(* IEC 61131-3 sources: SortJet_MasterSPS_Aufbau.fbsproj/09_Station/Shuttle/Bewegung, 2 files *)

(* ---- Querfahrt_Shuttle_FB_V01_00_00.fb.st ---- *)
(* METADATA
{
	"v3Meta": {
		"objectGuid": "72dffa9c-0dea-4fd7-9820-5307a69ebe3d"
	}
}
*)
FUNCTION_BLOCK Querfahrt_Shuttle_FB_V01_00_00
VAR_INPUT

  // BOOLEAN
  bpAktivieren                           : BOOL; // Hinweis: Baustein aktivieren
  bpReset                                : BOOL; // BETRIEBSART: Fehler zuruecksetzen
  bpReferenz                        : BOOL;
  bpHandfahrenPlus                             : BOOL;
  bpHandfahrenMinus                            : BOOL;
  bpFreigabe                             : BOOL; // Sicherheitsfreigabe Regler darf Freigeben
  bpAutomatikAktiv                       : BOOL; // BETRIEBSART: Umschaltung der Geschwindigkeit
  bpVerfahreShuttle                      : BOOL; // Befehl zum Positionieren
  bpVerfahrfreigabe                      : BOOL; // Das entsprechende Shutte setzt die Verfahrfreigabe und überträgt es an die Verfahrkontrolle
  bpSofortStop                           : BOOL;
  bpQuittungAuftragsstatusZurueckgesetzt : BOOL; // Auftrag wurde zurueckgesetzt
  bpTeilnehmerErreichbar                 : BOOL;
  bpShuttleFaecherwagenSuche             : BOOL;
  bpLangsamfahrtNockenAktivieren         : BOOL;

  // WORD
  wpAuftragsTyp                          : WORD; // Bit 1 = Positionierauftrag mit Messgeschwindigkeit (RackSuche), aus dem Positionierauftrag (Vorabpositionierung)

  // REAL
  rpDestinationPosition                  : REAL; // ZielPosition
  rpMinPosSwEsEingrenzung                : REAL;
  rpMaxPosSwEsEingrenzung                : REAL;

  // POINTER
  ppAntriebsInformationen  : REFERENCE TO AntriebsInformationen; // Hinweis: Beinhaltet die Geschwindigkeiten / Rampen der einzelnen Shuttle

  // STRUKTUR
  stStationsNummern     : Station_ST;

END_VAR
VAR_OUTPUT

  // BOOLEAN
  bpDone                         : BOOL;
  bpFehler                       : BOOL;
  bpPositionierungAktiv          : BOOL;
  bpAntriebLaeuft                : BOOL;
  bpInReference                  : BOOL;
  bpAuftragsstatusZuruecksetzen  : BOOL := FALSE;
  bpAbbruchPositionierung        : BOOL := FALSE;

  // WORD
  wpFehlerNr     : Fehlerkonstanten_EN; // Exception- Handle: Fehlernummer

  // REAL
  rpAktPosition : REAL;
  rpAktSpeed    : REAL;

  // HARDWARE EINGAENGE
  in_bLeistungsschutzFremdluefter : BOOL;
  in_bEndschalterMax              : BOOL; // Oeffner (TRUE = frei), gemappt; zum Umrichter ueber Signal-Steuerwort Bit 9, wirkt nur bei Endschalterquelle SPS
  in_bEndschalterMin              : BOOL; // Oeffner (TRUE = frei), gemappt; zum Umrichter ueber Signal-Steuerwort Bit 10, wirkt nur bei Endschalterquelle SPS

END_VAR
VAR

  // BOOLEAN
  Antrieb : REFERENCE TO Rexroth_ctrlX_Drive_Eckelmann_MC_V01_02_02;

  // BOOLEAN
  blErsterZyklus                : BOOL := TRUE;
  blFreigabeGesetzt             : BOOL;
  blAlterStatus_Bewegung        : BOOL;

  // REAL
  rlAlterStatus_Position        : REAL;

  // STEPS
  STEP_Mov_Shuttle_W    : Steps_TE;
  schrittlReset         : STEPS_TE;
  steplReferenz         : STEPS_TE;

  // TIMER
  tonlWarteAufStop                      : TON; // EINSCHALTVERZOEGERUNG:
  tonlWarteAufReset                     : TON; // EINSCHALTVERZOEGERUNG:
  tofAntriebFreigabe                    : TOF; // AUSSCHALTVERZÖGERUNG
  tonlEndschalterFreifahren             : TON;
  tonlWarteSchrittEndschalterFreifahren : TON;
  toflHardwareEndschalterFrei           : TOF;
  tonlSafetyTimeout                     : TON;
  tonlFreigabe                          : TON;
  tonlAntriebNichtBetriebsbereit        : TON;
  tonlStatusMelden                      : TON;

  // TRIGGER
  rtlAutoAktiv : R_TRIG;

END_VAR

//-------------------------------------------------------------------------------------------------
// S T A R T - Initialisierung
//-------------------------------------------------------------------------------------------------
IF ( blErsterZyklus ) THEN

  IF ( __ISVALIDREF(ppAntriebsInformationen) ) THEN

    blErsterZyklus := FALSE;

    Antrieb REF= pgAntriebe[ppAntriebsInformationen.wAchsID];

    (* Hinweis:
       - Initialisierung Antriebsinformationen
    *)
    Antrieb.ppAntriebsInformationen REF= ppAntriebsInformationen;
    Antrieb.stStationsNummern := stStationsNummern;

    (* Hinweis:
       - Für die Zielpunktkontrolle muss im ersten Zyklus (und nach jeder Referenzierung) die Zielposition initialisiert werden
    *)
    Antrieb.rpZielPosition := Antrieb.rpIstPosition;

    (* Hinweis:
       - Antriebswerte vorinitialisieren
    *)
    Antrieb.rpGeschwindigkeit := ppAntriebsInformationen.rpHandGeschwindigkeit;
    Antrieb.rpBeschleunigung  := ppAntriebsInformationen.rpMaxBeschleunigung;
    Antrieb.rpVerzoegerung    := ppAntriebsInformationen.rpMaxVerzoegerung;
    Antrieb.rpRuckzeit        := ppAntriebsInformationen.rpMaxRuckzeit;

  ELSE
    RETURN;
  END_IF

END_IF

//-------------------------------------------------------------------------------------------------
// E N D E - Initialisierung
//-------------------------------------------------------------------------------------------------

// Endschalter zyklisch an den Antrieb geben, auch bei deaktivierter Bewegung
Antrieb.bpEndschalterMinExtern := in_bEndschalterMin;
Antrieb.bpEndschalterMaxExtern := in_bEndschalterMax;

//-------------------------------------------------------------------------------------------------
// DEAKTIVIEREN
//-------------------------------------------------------------------------------------------------
IF ( NOT bpAktivieren ) THEN

  bpDone                        := TRUE;
  bpAuftragsstatusZuruecksetzen := FALSE;
  bpAbbruchPositionierung       := FALSE;

  bpFehler   := FALSE;
  wpFehlerNr := cMELDUNG_NULL;

  Antrieb.bpFreigabe := FALSE;

  RETURN;

END_IF

//-------------------------------------------------------------------------------------------------
// S T A R T - Timer
//-------------------------------------------------------------------------------------------------

rtlAutoAktiv(CLK := bpAutomatikAktiv);

IF ( rtlAutoAktiv.Q ) THEN
  Antrieb.rpZielPosition := Antrieb.rpIstPosition;
END_IF

(* Hinweis:
   - Aktuell wird diese Einschaltverzoegerung nur bei Motoren mit Bremse benoetigt [Lenze]
     => Eingebunden bei den Handfunktionen
*)
tofAntriebFreigabe( IN := blFreigabeGesetzt AND Antrieb.bpReglerBereit  , PT := T#10S );

// *************************************************************************************************

//-------------------------------------------------------------------------------------------------
// S T A R T - Verfahrschrittketten zurücksetzen
//-------------------------------------------------------------------------------------------------

// *************************************************************************************************

IF (   bpVerfahrfreigabe
     AND bpAbbruchPositionierung
     AND bpQuittungAuftragsstatusZurueckgesetzt )
THEN
  bpAbbruchPositionierung := FALSE;
  bpAuftragsstatusZuruecksetzen := FALSE;
  bpQuittungAuftragsstatusZurueckgesetzt := FALSE;

  wSps2MmiStationsNummer     := stStationsNummern.NummerIntern;
  rSps2MmiPosition           := Antrieb.rpIstPosition;
  MsgToMmi(SB0_SPS_SHUTTLEVORABPOSITIONIERUNGREADY);

END_IF

//-------------------------------------------------------------------------------------------------
// S T A R T - BAUSTEINE AUFRUFEN
//-------------------------------------------------------------------------------------------------

//-------------------------------------------------------------------------------------------------
// S T A R T - BAUSTEINE AUFRUFEN
//-------------------------------------------------------------------------------------------------
Verfahren();
Handfunktionen();
Referenz();
Reset();
Meldungen();

//-------------------------------------------------------------------------------------------------
// E N D E - BAUSTEINE AUFRUFEN
//-------------------------------------------------------------------------------------------------
IF ( bpSofortStop OR NOT abgVerfahrfreigabeShuttle[stStationsNummern.NummerSPS] ) OR NOT bpFreigabe THEN
  Antrieb.bpFreigabe := FALSE;
END_IF

Antrieb.stStationsNummern            := stStationsNummern;

Antrieb.bpAktiviereLangsamfahrtNocke := bpLangsamfahrtNockenAktivieren;
Antrieb.rpMinSwEsEingrenzung         := rpMinPosSwEsEingrenzung;
Antrieb.rpMaxSwEsEingrenzung         := rpMaxPosSwEsEingrenzung;

// übergabe der aktuellen Position
rpAktPosition   := Antrieb.rpIstPosition;
rpAktSpeed      := Antrieb.rpIstGeschwindigkeit; // mm/s, mit Vorzeichen
bpInReference   := Antrieb.bpIstReferenziert;
bpAntriebLaeuft := Antrieb.bpAntrieblaeuft;

// STATUS AN MMI MELDEN
tonlStatusMelden(
                  IN := NOT tonlStatusMelden.Q,
                  PT := T#500MS
                );

// Neue MMI-Verbindung (Flanke, nur ein Zyklus) sofort melden, nicht nur im 500-ms-Takt
IF    (     tonlStatusMelden.Q
        AND (    ( ABS( Antrieb.rpIstPosition - rlAlterStatus_Position ) > 1.0 )
              OR ( Antrieb.bpAntrieblaeuft <> blAlterStatus_Bewegung ) ) )
   OR Job.rtlMmiOk.Q
THEN
  stStationUpdate.wStationsNummer       := stStationsNummern.NummerSPS;
  stStationUpdate.eUpdateTyp            := StationUpdateTyp_EN.POSITIONSAENDERUNG;
  stStationUpdate.wAnzahlWerte          := 2;
  stStationUpdate.astWerte[1].eDatenTyp := UpdateDatenTyp_EN.TYP_REAL;
  stStationUpdate.astWerte[1].rWert     := Antrieb.rpIstPosition;
  stStationUpdate.astWerte[2].eDatenTyp := UpdateDatenTyp_EN.TYP_BOOL;
  stStationUpdate.astWerte[2].bWert     := Antrieb.bpAntrieblaeuft;
  MsgToMmi( auftragsnr_w := SB0_SPS_STATION_UPDATE );

  rlAlterStatus_Position := Antrieb.rpIstPosition;
  blAlterStatus_Bewegung := Antrieb.bpAntrieblaeuft;
END_IF
END_FUNCTION_BLOCK

(* ---- Verfahrueberwachung_PRG.prg.st ---- *)
(* METADATA
{
	"v3Meta": {
		"objectGuid": "88539335-6d2a-4efd-8213-a5feda61f359"
	}
}
*)
PROGRAM Verfahrueberwachung_PRG
VAR

  // BOOLEAN
  ablKonfiguriert                           : ARRAY[cERSTES_SHUTTLE..cLETZTES_TRANSFERSHUTTLE] OF BOOL; // Shuttle / Transfershuttle ist in dieser Anlage vorhanden
  ablShuttleInParkpos                       : ARRAY[cERSTES_SHUTTLE..cLETZTES_TRANSFERSHUTTLE] OF BOOL;
  ablShuttleStehtOhnePositionsveraenderung  : ARRAY[cERSTES_SHUTTLE..cLETZTES_TRANSFERSHUTTLE] OF BOOL;
  ablInReferenz                             : ARRAY[cERSTES_SHUTTLE..cLETZTES_TRANSFERSHUTTLE] OF BOOL; // Querfahrt-Antrieb referenziert (direkt aus pgAntriebe)

  // WORD
  wlIndex    : WORD;
  wlAchsID   : WORD; // Achs-ID des Querfahrt-Antriebs

  // REAL
  rlAlteZeit                               : REAL;
  rlAktuelleZeit                           : REAL;
  rlZyklusZeit                             : REAL;
  arlAktuelleGeschwindigkeit               : ARRAY[cERSTES_SHUTTLE..cLETZTES_TRANSFERSHUTTLE] OF REAL; // mm/s
  arlErrechneteGeschwindigkeit             : ARRAY[cERSTES_SHUTTLE..cLETZTES_TRANSFERSHUTTLE] OF REAL; // mm/s, aus der Positionsaenderung
  arlBerechneterBremsWeg                   : ARRAY[cERSTES_SHUTTLE..cLETZTES_TRANSFERSHUTTLE] OF REAL;
  arlAltePosition                          : ARRAY[cERSTES_SHUTTLE..cLETZTES_TRANSFERSHUTTLE] OF REAL;
  arlNeuePosition                          : ARRAY[cERSTES_SHUTTLE..cLETZTES_TRANSFERSHUTTLE] OF REAL;
  arlPostionsveraenderung                  : ARRAY[cERSTES_SHUTTLE..cLETZTES_TRANSFERSHUTTLE] OF REAL;
  arlErrechneteStillstandposition          : ARRAY[cERSTES_SHUTTLE..cLETZTES_TRANSFERSHUTTLE] OF REAL;
  arlVerzoegerung                          : ARRAY[cERSTES_SHUTTLE..cLETZTES_TRANSFERSHUTTLE] OF REAL; // Verzoegerung bei Sofort-Stopp in mm/s^2
  arlBremsfaktor                           : ARRAY[cERSTES_SHUTTLE..cLETZTES_TRANSFERSHUTTLE] OF REAL; // Bremszeit in s
  arlAktuellerSicherheitsabstand           : ARRAY[cERSTES_SHUTTLE..cLETZTES_TRANSFERSHUTTLE] OF REAL;
  arlPostionsMittelwert                    : ARRAY[cERSTES_SHUTTLE..cLETZTES_TRANSFERSHUTTLE] OF REAL;
  arlActPosShuttle                         : ARRAY[cERSTES_SHUTTLE..cLETZTES_TRANSFERSHUTTLE] OF REAL; // Aktuelle Position in mm
  arlActGeschwindigkeit                    : ARRAY[cERSTES_SHUTTLE..cLETZTES_TRANSFERSHUTTLE] OF REAL; // Aktuelle Geschwindigkeit in mm/s

  // STRUCT
  arrParkpositionen                        : ARRAY[cERSTES_SHUTTLE..cLETZTES_TRANSFERSHUTTLE] OF Parkpositionen_ST;

  // TIME
  TmStmp : TIME;
  Zyklus : TIME;

END_VAR
VAR CONSTANT

  // REAL
  cTOLERANZ_PARKPOSITION : REAL := 100.0; // Abweichung zur Parkposition [mm], in der das Shuttle als "in Parkposition" gilt
  cTOLERANZ_STEHT        : REAL := 2.0;   // Positionsaenderung je Zyklus [mm], unter der das Shuttle als stehend gilt

END_VAR
(* Hinweis:
   - Dieser Baustein errechnet die Stillstandsposition von fahrenden Shuttlen (Shuttle und Transfershuttle),
     um eine drohende Kollision zweier Shuttle auf einer Bahn vorauszuberechnen.
   - Die berechneten Einheiten sind mm und s.
   - Die Shuttle liegen auf einer Bahn in der Reihenfolge ihrer Nummer: das Shuttle mit der kleineren Nummer
     (z. B. 151) liegt auf der kleineren Position, das mit der groesseren Nummer (z. B. 152) auf der groesseren.
*)
TmStmp := TIME();

//-------------------------------------------------------------------------------------------------
// BAUSTEIN: ZYKLUSZEITBERECHNUNG
//-------------------------------------------------------------------------------------------------
rlAktuelleZeit := TIME_TO_REAL(TIME());
rlZyklusZeit   := rlAktuelleZeit - rlAlteZeit;
rlAlteZeit     := rlAktuelleZeit;

// WORKAROUND EXCEPTION
IF ( rlZyklusZeit = 0 ) THEN
  rlZyklusZeit := 1;
END_IF

//-------------------------------------------------------------------------------------------------
// BAUSTEIN: UEBERGABE PARKPOSITION, VERZOEGERUNG UND POSITION
//-------------------------------------------------------------------------------------------------
(* Hinweis:
   - Parkpositionen, Verzoegerungen (Maschinenkonstanten, in mm/s^2) und die vom Antrieb gemeldete Position / Geschwindigkeit
     der Shuttle und der Transfershuttle in gemeinsame Arrays uebernehmen
   - Ist ein Shuttle deaktiviert, wird seine Position auf die weit entfernte Parkseite gelegt, damit es nicht stoert
*)
FOR wlIndex := cERSTES_SHUTTLE TO cLETZTES_SHUTTLE DO

  IF NOT __ISVALIDREF(starrShuttleBasisParameter[wlIndex].stMKs) THEN
    abgVerfahrfreigabeShuttle[wlIndex] := FALSE;
    ablKonfiguriert[wlIndex] := FALSE;
    CONTINUE;
  END_IF

  ablKonfiguriert[wlIndex] := ( apgShuttleVerfahrparameter[wlIndex].eParkposition = PARKPOSITION_MAX
                                OR apgShuttleVerfahrparameter[wlIndex].eParkposition = PARKPOSITION_MIN
                                OR apgShuttleVerfahrparameter[wlIndex].eParkposition = PARKPOSITION_MIN_MAX );

  IF ablKonfiguriert[wlIndex] THEN

    arrParkpositionen[wlIndex].eParkposition        := apgShuttleVerfahrparameter[wlIndex].eParkposition;
    arrParkpositionen[wlIndex].rParkpositionMaximum := apgShuttleVerfahrparameter[wlIndex].rParkpositionMaximum;
    arrParkpositionen[wlIndex].rParkpositionMinimum := apgShuttleVerfahrparameter[wlIndex].rParkpositionMinimum;
    arlVerzoegerung[wlIndex]                        := apgVerfahrueberwachung[wlIndex].rMaxVerzoegerungsRampeUeberwachung;

    (* Hinweis:
       - Position / Geschwindigkeit / Referenz direkt aus dem Querfahrt-Antrieb (pgAntriebe, laeuft ebenfalls in der FastTask)
       - NICHT ueber aShuttle[].Querfahrt lesen: das ist eine Instanz der MainTask -> Mehrfach-Task-Zugriff auf deren E/As (C0373)
    *)
    IF (     NOT starrShuttleBasisParameter[wlIndex].stMKs.bDeaktivieren
         AND __ISVALIDREF(starrShuttleBasisParameter[wlIndex].stAntriebsparameter.stQuerfahrt) )
    THEN
      wlAchsID                       := starrShuttleBasisParameter[wlIndex].stAntriebsparameter.stQuerfahrt.wAchsID;
      arlActPosShuttle[wlIndex]      := pgAntriebe[wlAchsID].rpIstPosition;
      arlActGeschwindigkeit[wlIndex] := pgAntriebe[wlAchsID].rpIstGeschwindigkeit;
      ablInReferenz[wlIndex]         := pgAntriebe[wlAchsID].bpIstReferenziert;
    ELSE
      arlActPosShuttle[wlIndex]      := SEL( apgShuttleVerfahrparameter[wlIndex].eParkposition = PARKPOSITION_MAX, -50000.0, 50000.0 );
      arlActGeschwindigkeit[wlIndex] := 0;
      ablInReferenz[wlIndex]         := FALSE;
    END_IF

  ELSE
    wpgFehlerdaten[0] := wlIndex;
    wpgFehlerdaten[1] := apgShuttleVerfahrparameter[wlIndex].eParkposition;
    SpsHinweis( eFehler_Verfahrueberwachung,
                cMELDUNG_VERFAHRUEBERWACHUNG_UNGUELTIGE_PARKPOSITION,
                wlIndex,
                AutomatikkreisBestimmen(wlIndex),
                wpgFehlerdaten );
  END_IF

END_FOR

FOR wlIndex := cERSTES_TRANSFERSHUTTLE TO cLETZTES_TRANSFERSHUTTLE DO

  IF NOT __ISVALIDREF(starrTransfershuttleBasisParameter[wlIndex].stMKs) THEN
    abgVerfahrfreigabeShuttle[wlIndex] := FALSE;
    ablKonfiguriert[wlIndex] := FALSE;
    CONTINUE;
  END_IF

  ablKonfiguriert[wlIndex] := ( apgTransfershuttleVerfahrparameter[wlIndex].eParkposition = PARKPOSITION_MAX
                                OR apgTransfershuttleVerfahrparameter[wlIndex].eParkposition = PARKPOSITION_MIN
                                OR apgTransfershuttleVerfahrparameter[wlIndex].eParkposition = PARKPOSITION_MIN_MAX );

  IF ablKonfiguriert[wlIndex] THEN

    arrParkpositionen[wlIndex].eParkposition        := apgTransfershuttleVerfahrparameter[wlIndex].eParkposition;
    arrParkpositionen[wlIndex].rParkpositionMaximum := apgTransfershuttleVerfahrparameter[wlIndex].rParkpositionMaximum;
    arrParkpositionen[wlIndex].rParkpositionMinimum := apgTransfershuttleVerfahrparameter[wlIndex].rParkpositionMinimum;
    arlVerzoegerung[wlIndex]                        := apgVerfahrueberwachungTransfershuttle[wlIndex].rMaxVerzoegerungsRampeUeberwachung;

    (* Hinweis:
       - Position / Geschwindigkeit / Referenz direkt aus dem Querfahrt-Antrieb (pgAntriebe, laeuft ebenfalls in der FastTask)
       - NICHT ueber aTransfershuttles[].Querfahrt lesen: das ist eine Instanz der MainTask -> Mehrfach-Task-Zugriff auf deren E/As (C0373)
    *)
    IF (     NOT starrTransfershuttleBasisParameter[wlIndex].stMKs.bDeaktivieren
         AND __ISVALIDREF(starrTransfershuttleBasisParameter[wlIndex].stAntriebsparameter.stQuerfahrt) )
    THEN
      wlAchsID                       := starrTransfershuttleBasisParameter[wlIndex].stAntriebsparameter.stQuerfahrt.wAchsID;
      arlActPosShuttle[wlIndex]      := pgAntriebe[wlAchsID].rpIstPosition;
      arlActGeschwindigkeit[wlIndex] := pgAntriebe[wlAchsID].rpIstGeschwindigkeit;
      ablInReferenz[wlIndex]         := pgAntriebe[wlAchsID].bpIstReferenziert;
    ELSE
      arlActPosShuttle[wlIndex]      := SEL( apgTransfershuttleVerfahrparameter[wlIndex].eParkposition = PARKPOSITION_MAX, -50000.0, 50000.0 );
      arlActGeschwindigkeit[wlIndex] := 0;
      ablInReferenz[wlIndex]         := FALSE;
    END_IF

  ELSE
    wpgFehlerdaten[0] := wlIndex;
    wpgFehlerdaten[1] := apgTransfershuttleVerfahrparameter[wlIndex].eParkposition;
    SpsHinweis( eFehler_Verfahrueberwachung,
                cMELDUNG_VERFAHRUEBERWACHUNG_UNGUELTIGE_PARKPOSITION,
                wlIndex,
                AutomatikkreisBestimmen(wlIndex),
                wpgFehlerdaten );
  END_IF

END_FOR

//-------------------------------------------------------------------------------------------------
// BAUSTEIN: STILLSTANDSPOSITION UND PARKPOSITION
//-------------------------------------------------------------------------------------------------
(* Hinweis:
   - Bei einem stillstehenden Shuttle ist die errechnete Stillstandsposition gleich der aktuellen Position
   - Sonst: Position plus Bremsweg bei Sofort-Stopp in Fahrtrichtung
*)
FOR wlIndex := cERSTES_SHUTTLE TO cLETZTES_TRANSFERSHUTTLE DO

  IF NOT ablKonfiguriert[wlIndex] THEN
    CONTINUE;
  END_IF

  // => Die alte Position minus der neuen Position ergibt die Positionsveraenderung,
  //      geteilt durch die Zykluszeit ergibt das Weg/Zeit -> mm/ms, mal 1000 ergibt mm/s
  arlNeuePosition[wlIndex]                          := arlActPosShuttle[wlIndex];
  arlPostionsveraenderung[wlIndex]                  := arlNeuePosition[wlIndex] - arlAltePosition[wlIndex];
  arlErrechneteGeschwindigkeit[wlIndex]             := ( arlPostionsveraenderung[wlIndex] / rlZyklusZeit ) * 1000;
  ablShuttleStehtOhnePositionsveraenderung[wlIndex] := ( ABS( arlPostionsveraenderung[wlIndex] ) < 1 );

  // Mittelwert aus alter und neuer Position, VOR dem Ueberschreiben der alten Position bilden
  arlPostionsMittelwert[wlIndex] := ( arlNeuePosition[wlIndex] + arlAltePosition[wlIndex] ) / 2;
  arlAltePosition[wlIndex]       := arlNeuePosition[wlIndex];

  arlAktuelleGeschwindigkeit[wlIndex] := arlActGeschwindigkeit[wlIndex]; // mm/s

  // => Verbleibende Wegstrecke bei einem Sofort-Stopp
  //   => Berechnung:
  //      F [mm/s], a [mm/s^2], S [mm], t [s]
  //
  //      S = ( ( Va-Ve ) / 2 ) * t
  //      t = Va / a
  //
  //      S = ( ( Va-Ve ) / 2 ) * ( Va / a )
  //
  //      fuer Ve gilt = 0
  //
  //      S = ( Va / 2 ) * ( Va / a )
  IF ( arlVerzoegerung[wlIndex] > 0 ) THEN
    arlBremsfaktor[wlIndex] := arlAktuelleGeschwindigkeit[wlIndex] / arlVerzoegerung[wlIndex]; // dies ist t
  ELSE
    arlBremsfaktor[wlIndex] := 0;
  END_IF

  arlBerechneterBremsWeg[wlIndex] := ( arlAktuelleGeschwindigkeit[wlIndex] / 2.0 ) * arlBremsfaktor[wlIndex];

  // => Der errechnete Bremsweg ist durch die Quadratur immer positiv, deshalb nach Fahrtrichtung unterscheiden
  IF ( arlAktuelleGeschwindigkeit[wlIndex] > 0 ) THEN
    arlErrechneteStillstandposition[wlIndex] := arlNeuePosition[wlIndex] + arlBerechneterBremsWeg[wlIndex];
  ELSE
    arlErrechneteStillstandposition[wlIndex] := arlNeuePosition[wlIndex] - arlBerechneterBremsWeg[wlIndex];
  END_IF

  (* Hinweis:
     - Wenn das Shuttle in Parkposition ist, darf das Gegenshuttle naeher fahren
  *)
  CASE arrParkpositionen[wlIndex].eParkposition OF

    PARKPOSITION_MIN:
      ablShuttleInParkpos[wlIndex] :=
                                     ABS( arlErrechneteStillstandposition[wlIndex] - arrParkpositionen[wlIndex].rParkpositionMinimum ) < cTOLERANZ_PARKPOSITION // im Bereich der Parkposition
                                     AND ( ABS( arlPostionsMittelwert[wlIndex] - arlNeuePosition[wlIndex] ) < cTOLERANZ_STEHT ); // das Shuttle steht

    PARKPOSITION_MAX:
      ablShuttleInParkpos[wlIndex] :=
                                     ABS( arlErrechneteStillstandposition[wlIndex] - arrParkpositionen[wlIndex].rParkpositionMaximum ) < cTOLERANZ_PARKPOSITION // im Bereich der Parkposition
                                     AND ( ABS( arlPostionsMittelwert[wlIndex] - arlNeuePosition[wlIndex] ) < cTOLERANZ_STEHT ); // das Shuttle steht

    PARKPOSITION_MIN_MAX:
      ablShuttleInParkpos[wlIndex] :=
                                     (
                                       ( ABS( arlErrechneteStillstandposition[wlIndex] - arrParkpositionen[wlIndex].rParkpositionMinimum ) < cTOLERANZ_PARKPOSITION )
                                       OR ( ABS( arlErrechneteStillstandposition[wlIndex] - arrParkpositionen[wlIndex].rParkpositionMaximum ) < cTOLERANZ_PARKPOSITION )
                                     ) // im Bereich der Parkposition
                                     AND ( ABS( arlPostionsMittelwert[wlIndex] - arlNeuePosition[wlIndex] ) < cTOLERANZ_STEHT ); // das Shuttle steht

  END_CASE

END_FOR

//-------------------------------------------------------------------------------------------------
// BAUSTEIN: ABSTANDSUEBERWACHUNG TRANSFERSHUTTLE 151 <-> 152
//-------------------------------------------------------------------------------------------------
(* Hinweis:
   - Die Transfershuttle 151 und 152 fahren auf einer Bahn, 151 liegt auf der kleineren Position
   - Ist eines der beiden in Parkposition, gilt der kleinere Abstand
   - Die Verfahrfreigabe wird jeden Zyklus neu gebildet und nur gesperrt, solange der Mindestabstand unterschritten wuerde
   - Gesperrt wird nur, wenn beide Transfershuttle referenziert sind
*)
IF ( ablShuttleInParkpos[cSHUTTLE_151] OR ablShuttleInParkpos[cSHUTTLE_152] ) THEN
  arlAktuellerSicherheitsabstand[cSHUTTLE_151] := rgMkMinSecureDistanceTransferAtParkPos;
  arlAktuellerSicherheitsabstand[cSHUTTLE_152] := rgMkMinSecureDistanceTransferAtParkPos;
ELSE
  arlAktuellerSicherheitsabstand[cSHUTTLE_151] := rgMkMinSecureDistanceTransfer;
  arlAktuellerSicherheitsabstand[cSHUTTLE_152] := rgMkMinSecureDistanceTransfer;
END_IF

abgVerfahrfreigabeShuttle[cSHUTTLE_151] := __ISVALIDREF(starrTransfershuttleBasisParameter[cSHUTTLE_151].stMKs);
abgVerfahrfreigabeShuttle[cSHUTTLE_152] := __ISVALIDREF(starrTransfershuttleBasisParameter[cSHUTTLE_152].stMKs);

IF ablInReferenz[cSHUTTLE_151]
   AND ablInReferenz[cSHUTTLE_152]
THEN

  // 151 darf nicht ueber 152 hinaus (minus Sicherheitsabstand)
  IF arlErrechneteStillstandposition[cSHUTTLE_151] >
     ( arlErrechneteStillstandposition[cSHUTTLE_152] - arlAktuellerSicherheitsabstand[cSHUTTLE_151] )
  THEN
    abgVerfahrfreigabeShuttle[cSHUTTLE_151] := FALSE;
  END_IF

  // 152 darf nicht unter 151 hinaus (plus Sicherheitsabstand)
  IF arlErrechneteStillstandposition[cSHUTTLE_152] <
     ( arlErrechneteStillstandposition[cSHUTTLE_151] + arlAktuellerSicherheitsabstand[cSHUTTLE_152] )
  THEN
    abgVerfahrfreigabeShuttle[cSHUTTLE_152] := FALSE;
  END_IF

END_IF

//-------------------------------------------------------------------------------------------------
// BAUSTEIN: ABSTANDSUEBERWACHUNG SHUTTLE 101 <-> 102 (DUMMY, AUSKOMMENTIERT)
//-------------------------------------------------------------------------------------------------
(* Hinweis:
   - Nur noetig, wenn sich zwei Shuttle auf EINER Bahn befinden (bei getrennten Bahnen nicht: 101 und 102 fahren dann unabhaengig)
   - Zum Aktivieren: Kommentar entfernen. MKs rgMkMinSecureDistanceShuttles / ...AtParkPos sind vorhanden
   - Aufbau wie bei den Transfershuttle: 101 liegt auf der kleineren Position, 102 auf der groesseren
   - Fuer weitere Paare auf einer Bahn kopieren und die Nummern anpassen

     IF ( ablShuttleInParkpos[cSHUTTLE_101] OR ablShuttleInParkpos[cSHUTTLE_102] ) THEN
     arlAktuellerSicherheitsabstand[cSHUTTLE_101] := rgMkMinSecureDistanceShuttlesAtParkPos;
     arlAktuellerSicherheitsabstand[cSHUTTLE_102] := rgMkMinSecureDistanceShuttlesAtParkPos;
     ELSE
     arlAktuellerSicherheitsabstand[cSHUTTLE_101] := rgMkMinSecureDistanceShuttles;
     arlAktuellerSicherheitsabstand[cSHUTTLE_102] := rgMkMinSecureDistanceShuttles;
     END_IF

     abgVerfahrfreigabeShuttle[cSHUTTLE_101] := TRUE;
     abgVerfahrfreigabeShuttle[cSHUTTLE_102] := TRUE;

     IF ablInReferenz[cSHUTTLE_101]
     AND ablInReferenz[cSHUTTLE_102]
     THEN

     IF arlErrechneteStillstandposition[cSHUTTLE_101] >
     ( arlErrechneteStillstandposition[cSHUTTLE_102] - arlAktuellerSicherheitsabstand[cSHUTTLE_101] )
     THEN
     abgVerfahrfreigabeShuttle[cSHUTTLE_101] := FALSE;
     END_IF

     IF arlErrechneteStillstandposition[cSHUTTLE_102] <
     ( arlErrechneteStillstandposition[cSHUTTLE_101] + arlAktuellerSicherheitsabstand[cSHUTTLE_102] )
     THEN
     abgVerfahrfreigabeShuttle[cSHUTTLE_102] := FALSE;
     END_IF

     END_IF
*)

Zyklus := TIME() - TmStmp;
END_PROGRAM
